{region 'Documentation'}
(*!
<summary>Thin TestSuiteBase subject with a typed child array and isolated dependencies.</summary>
<description>
Bind is called before Initialize. Production initialization, sequencing, aggregation and
publication remain inherited. Configure records its context and builds a small real collection.
The uninitialized-child option uses a separate never-initialized double, not mutated base state.
ProcessTestCases applies the scenario's child view only after the base has called its helper.
</description>
*)
{endregion}
FUNCTION_BLOCK TestSuiteLifecycleProbe EXTENDS TestSuiteBase
VAR
    FChildA : SuiteLifecycleChildDouble;
    FChildB : SuiteLifecycleChildDouble;
    FUninitializedChild : SuiteLifecycleChildDouble;
    FTestCases : ARRAY[4..6] OF I_TestCase;
    FChildObservation : ST_OrchestrationObservation;
    FSecondChildObservation : ST_OrchestrationObservation;
    FRegisterChildren : BOOL := TRUE;
    FIncludeUninitializedChild : BOOL;
    FConfigureCount : UINT;
    FConfigureContextValid : BOOL;
    FChildCallCount : UINT;
END_VAR

SUPER^();

{region 'Documentation'}
(*!
<summary>Binds isolated dependencies before Initialize and selects the concrete setup to exercise.</summary>
*)
{endregion}
METHOD PUBLIC Bind
VAR_INPUT
    Publisher : I_EventPublisher; //! Nonzero isolated event publisher retained before subject initialization; keep it alive through all subject use.
    Helper : I_Orchestrator; //! Nonzero injected orchestration helper retained before owner initialization; keep it alive through subject use.
    RegisterChildren : BOOL := TRUE; //! TRUE registers the two controlled children; FALSE exercises empty configuration.
    IncludeUninitializedChild : BOOL := FALSE; //! TRUE leaves a registered controlled child uninitialized to exercise rejection.
END_VAR
FEventPublisher := Publisher;
FOrchestrator := Helper;
FRegisterChildren := RegisterChildren;
FIncludeUninitializedChild := IncludeUninitializedChild;
FChildA.SetReleaseResponse();
FChildB.SetReleaseResponse();
FConfigureCount := 0;
FChildCallCount := 0;
FConfigureContextValid := FALSE;
FChildObservation.State := E_State.Uninitialized;
FChildObservation.Result := E_Result.NotEvaluated;
FChildObservation.Ready := FALSE;
FChildObservation.Complete := FALSE;
FSecondChildObservation := FChildObservation;
END_METHOD

{region 'Documentation'}
(*!
<summary>Both concrete child bodies have executed exactly once per ProcessTestCases invocation.</summary>
*)
{endregion}
{attribute 'monitoring' := 'call'}
PROPERTY PUBLIC ChildBodyCallsMatch : BOOL //! Both concrete child bodies have executed exactly once per ProcessTestCases invocation.
GET
VAR
    FirstCalls : ST_OrchestrationCalls;
    SecondCalls : ST_OrchestrationCalls;
END_VAR
FirstCalls := FChildA.Calls;
SecondCalls := FChildB.Calls;
ChildBodyCallsMatch := (FirstCalls.BodyCount = FChildCallCount) AND (SecondCalls.BodyCount = FChildCallCount);
END_GET
END_PROPERTY

{region 'Documentation'}
(*!
<summary>Number of ProcessTestCases invocations since binding.</summary>
*)
{endregion}
{attribute 'monitoring' := 'call'}
PROPERTY PUBLIC ChildCallCount : UINT //! Number of ProcessTestCases invocations since binding.
GET
ChildCallCount := FChildCallCount;
END_GET
END_PROPERTY

{region 'Documentation'}
(*!
<summary>Registers two controlled typed children in a shifted array with spare capacity; records base context.</summary>
*)
{endregion}
METHOD PROTECTED Configure
VAR_IN_OUT
    // SA0167: Borrowed setup builder; no temporary instance is created.
    {attribute 'analysis' := '-167'}
    Builder : TestSuiteConfigurationBuilder; //! Borrowed owner configuration builder used only during this Configure call; register this owner's concrete children.
END_VAR
FConfigureCount := FConfigureCount + 1;
FConfigureContextValid := (State = E_State.Uninitialized) AND NOT IsInitialized AND (Name <> '');
Builder.Initialize(Mode := E_OrchestrationMode.Serial,
    TestCases := FTestCases);
FChildA.Initialize(Name := CONCAT(Name, '.ChildA'),
    Slot := 0);
FChildB.Initialize(Name := CONCAT(Name, '.ChildB'),
    Slot := 0);
IF NOT FRegisterChildren THEN
    RETURN;
END_IF;
Builder.Register(TestCase := FChildA);
IF FIncludeUninitializedChild THEN
    Builder.Register(TestCase := FUninitializedChild);
ELSE
    Builder.Register(TestCase := FChildB);
END_IF;
END_METHOD

{region 'Documentation'}
(*!
<summary>Configure saw the new identity before successful initialization.</summary>
*)
{endregion}
{attribute 'monitoring' := 'call'}
PROPERTY PUBLIC ConfigureContextValid : BOOL //! Configure saw the new identity before successful initialization.
GET
ConfigureContextValid := FConfigureContextValid;
END_GET
END_PROPERTY

{region 'Documentation'}
(*!
<summary>Number of Configure calls since binding.</summary>
*)
{endregion}
{attribute 'monitoring' := 'call'}
PROPERTY PUBLIC ConfigureCount : UINT //! Number of Configure calls since binding.
GET
ConfigureCount := FConfigureCount;
END_GET
END_PROPERTY

{region 'Documentation'}
(*!
<summary>Returns the recorded calls of a registered controlled child; unknown indices return an empty observation.</summary>
*)
{endregion}
METHOD PUBLIC GetChildCalls : ST_OrchestrationCalls //! Retained call trace for the selected child; an empty trace for an unknown index or empty collection.
VAR_INPUT
    Index : DINT; //! Original occupied child-array index; unknown indices return an empty trace.
END_VAR
VAR
    EmptyCalls : ST_OrchestrationCalls;
END_VAR
GetChildCalls := EmptyCalls;
IF ChildCount = 0 THEN
    RETURN;
END_IF;
IF Index = ChildArrayLowerBound THEN
    GetChildCalls := FChildA.Calls;
ELSIF (ChildCount > 1) AND (Index = ChildArrayLowerBound + 1) THEN
    GetChildCalls := FChildB.Calls;
END_IF;
END_METHOD

{region 'Documentation'}
(*!
<summary>Returns the registered typed entry by actual array index; lookup never executes a child.</summary>
*)
{endregion}
METHOD PUBLIC GetTestCase : I_TestCase //! Typed child interface at the original array index; zero when no entry is available.
VAR_INPUT
    Index : DINT; //! Original occupied child-array index, rather than an ordinal position.
END_VAR
GetTestCase := 0;
IF (ChildCount = 0) OR (Index < ChildArrayLowerBound)
    OR (DINT_TO_LINT(Index) >= DINT_TO_LINT(ChildArrayLowerBound) + UINT_TO_LINT(ChildCount)) THEN
    RETURN;
END_IF;
GetTestCase := FTestCases[Index];
END_METHOD

{region 'Documentation'}
(*!
<summary>Applies the next scripted observation after the helper; counts calls without replacing owner processing.</summary>
*)
{endregion}
METHOD PROTECTED ProcessTestCases
FChildA(ObservationInput := FChildObservation);
FChildB(ObservationInput := FSecondChildObservation);
FChildCallCount := FChildCallCount + 1;
END_METHOD

{region 'Documentation'}
(*!
<summary>Selects the next child snapshot; it becomes visible only in ProcessTestCases, after helper execution.</summary>
*)
{endregion}
METHOD PUBLIC SetChildObservation
VAR_INPUT
    Observation : ST_OrchestrationObservation; //! Scripted view copied to both children for acceptance on their next concrete body calls.
END_VAR
FChildObservation := Observation;
FSecondChildObservation := Observation;
END_METHOD

{region 'Documentation'}
(*!
<summary>Supplies independent next snapshots; each child accepts its view only when the Suite calls its body.</summary>
*)
{endregion}
METHOD PUBLIC SetChildObservations
VAR_INPUT
    FirstChild : ST_OrchestrationObservation; //! Scripted view for the first child, accepted on its next concrete body call.
    SecondChild : ST_OrchestrationObservation; //! Scripted view for the second child, accepted on its next concrete body call.
END_VAR
FChildObservation := FirstChild;
FSecondChildObservation := SecondChild;
END_METHOD

{region 'Documentation'}
(*!
<summary>Controls only the child release boundary for delegation tests, without changing Suite accounting.</summary>
*)
{endregion}
METHOD PUBLIC SetChildReleaseResponses
VAR_INPUT
    FirstSucceeds : BOOL := TRUE; //! Release response installed in the first controlled child.
    SecondSucceeds : BOOL := TRUE; //! Release response installed in the second controlled child.
END_VAR
FChildA.SetReleaseResponse(Succeeds := FirstSucceeds);
FChildB.SetReleaseResponse(Succeeds := SecondSucceeds);
END_METHOD

END_FUNCTION_BLOCK

(* stored: Version 1.1.0.1
   POU TestSuiteLifecycleProbe: Id {1339857b-5a9a-449d-bf48-ba5fe9b390c2}, SpecialFunc None
   Folder Internal: Id {d548c392-2496-4357-bbef-6bfe9477e753}
   Method Bind: Id {9605a89f-f2db-476b-8f6e-0085dc959049}
   Property ChildBodyCallsMatch: Id {dbff5695-7453-497c-83dd-a070f1599c9c}
   Get Get: Id {d82d9e20-d9c7-400d-a12a-d81ac934fdf8}
   Property ChildCallCount: Id {49f458d4-d6f4-4732-a608-8b03e7b59f18}
   Get Get: Id {96d2f627-cf97-48fb-b6c1-79d4eef450c9}
   Method Configure: Id {fb535502-d727-4a1a-93bb-9614d0b00dc0}
   Property ConfigureContextValid: Id {5e0365f3-d2b9-4872-9e7c-2d226659ec90}
   Get Get: Id {bd8fc4cf-0353-4d4d-96f5-29634381d1f8}
   Property ConfigureCount: Id {b2baff1e-491d-4e44-84ab-eab1715c44bb}
   Get Get: Id {700e0ffe-626e-428c-9799-3f7504c5a83d}
   Method GetChildCalls: Id {05e58dcd-281a-408a-a0f4-373bae016987}
   Method GetTestCase: Id {75e2507a-9fa3-4b0a-83c5-5e2657fd1499}
   Method ProcessTestCases: Id {4a2e09f3-f245-4564-9345-6e3a12fca529}
   Method SetChildObservation: Id {0b2b13bb-de11-49d2-b493-8861f578f990}
   Method SetChildObservations: Id {2f7e846e-a703-4f3d-a22a-804758c912f4}
   Method SetChildReleaseResponses: Id {2596f085-faae-47f6-81f5-02b673fcc2fd} *)
